(*
This is *emphasized text*.

This is **strong text**.

This text is an example of ``inline literals``.
*)

FUNCTION_BLOCK FB_Libdoc_FontStyle
VAR_INPUT
    nVarA : INT;
    nVarB : INT;
END_VAR
VAR_OUTPUT
    nSum : INT;
END_VAR
VAR
END_VAR

END_FUNCTION_BLOCK

(* stored: Version 1.1.0.1, ProductVersion 3.1.4022.17
   POU FB_Libdoc_FontStyle: Id {07ca8705-e54e-421c-bfc6-aceeebfd7728}, SpecialFunc None *)
